ABB RAPID module: PgProg.mod

MODULE MainModule
GLOBAL VAR robtarget robpoint0= p:{{-640.584, 506.980, 371.534},{0.374108, 0.285846, 0.853660, -0.222712}}{cfg 0,0,0,0}{EJ 0.000000000,0.000000000,0.000000000,0.000000000,0.000000000,0.000000000}
GLOBAL VAR robtarget robpoint1= p:{{-607.850, 543.849, 363.215},{0.374108, 0.285846, 0.853660, -0.222712}}{cfg 0,0,0,0}{EJ 0.000000000,0.000000000,0.000000000,0.000000000,0.000000000,0.000000000}
GLOBAL VAR robtarget robpoint2= p:{{-602.951, 596.788, 316.595},{0.374108, 0.285846, 0.853660, -0.222712}}{cfg 0,0,0,0}{EJ 0.000000000,0.000000000,0.000000000,0.000000000,0.000000000,0.000000000}
GLOBAL VAR robtarget robpoint3= p:{{-663.517, 575.988, 286.611},{0.374108, 0.285846, 0.853660, -0.222712}}{cfg 0,0,0,0}{EJ 0.000000000,0.000000000,0.000000000,0.000000000,0.000000000,0.000000000}
GLOBAL VAR robtarget robpoint4= p:{{-650.861, 503.437, 361.399},{0.374108, 0.285846, 0.853660, -0.222712}}{cfg 0,0,0,0}{EJ 0.000000000,0.000000000,0.000000000,0.000000000,0.000000000,0.000000000}
GLOBAL VAR robtarget robpoint5= p:{{-640.584, 506.980, 371.534},{0.374108, 0.285846, 0.853660, -0.222712}}{cfg 0,0,0,0}{EJ 0.000000000,0.000000000,0.000000000,0.000000000,0.000000000,0.000000000}
GLOBAL VAR robtarget robpoint6= p:{{-607.850, 543.849, 363.215},{0.374108, 0.285846, 0.853660, -0.222712}}{cfg 0,0,0,0}{EJ 0.000000000,0.000000000,0.000000000,0.000000000,0.000000000,0.000000000}
GLOBAL VAR robtarget robpoint7= p:{{-353.026, -90.135, 331.702},{0.344329, 0.048056, 0.933073, -0.092215}}{cfg -1,0,-1,0}{EJ 0.000000000,0.000000000,0.000000000,0.000000000,0.000000000,0.000000000}

GLOBAL Proc main()
    wobj16.x = 1234.57
    wobj16.y = -98.765
    wobj16.z = 50.500
    wobj16.q1 = 0.965926
    wobj16.q2 = 0.000000
    wobj16.q3 = 0.000000
    wobj16.q4 = 0.258819
    tool03.x = 10.000
    tool03.y = 20.000
    tool03.z = 150.000
    tool03.q1 = 0.991445
    tool03.q2 = 0.130526
    tool03.q3 = 0.000000
    tool03.q4 = 0.000000
    MoveJ robpoint0,v250,z5,tool03,wobj16
    MoveL robpoint1,v250,z5,tool03,wobj16
    MoveC robpoint2,robpoint3,v250,z5,tool03,wobj16
    MoveL robpoint4,v100,z5,tool03,wobj16
    MoveL robpoint5,v100,z0,tool03,wobj16
    Wait 0.500
    TPWrite "Hello from postgen";
    SubProgram;
    CustomCode(42)
    ThreadProg
    SetDO D_OUT_1, 1;
    SetDO Valve, 0;
    SetDO D_OUT_3, 2.5;
    WaitDI D_IN_2, 1;
    WaitDI D_IN_4, 0, \MaxTime:=1.5;
    tool03.x = 0.000
    tool03.y = 0.000
    tool03.z = 200.000
    tool03.q1 = 1.000000
    tool03.q2 = 0.000000
    tool03.q3 = 0.000000
    tool03.q4 = 0.000000
    MoveJ robpoint6,v100,z0,tool03,wobj16
    MoveL robpoint7,v100,z0,tool03,wobj16
EndProc
EndModule
